PROGRAM PRG_Ladder
VAR
    bStart, bStop, bMotor, bButton, bClear, bLamp, bSkip, bRunning, bAlarm, bReady : BOOL;
    tonRun : TON;
    tElapsed : TIME;
END_VAR
VAR // added by the converter: edge detectors and wires of the graphical bodies
    _rt1 : R_TRIG;
END_VAR

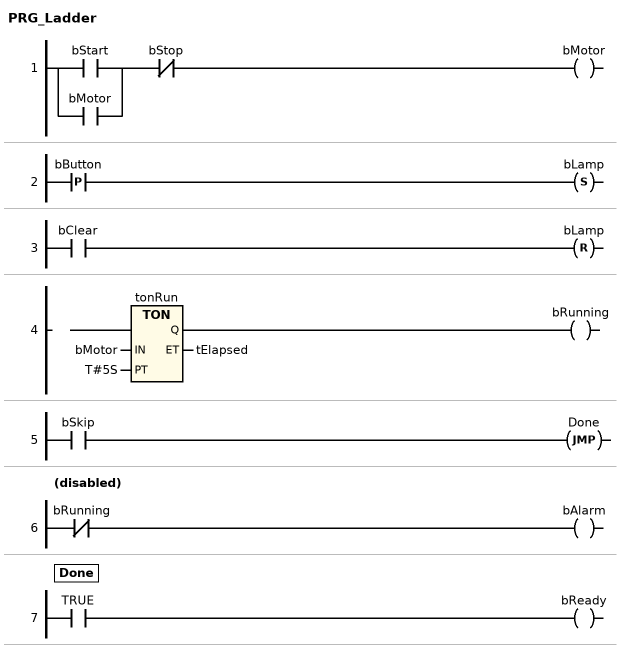
// NETWORK 1
bMotor := (bStart OR bMotor) AND NOT bStop;

// NETWORK 2
_rt1(CLK := bButton);
bLamp S= _rt1.Q;

// NETWORK 3
bLamp R= bClear;

// NETWORK 4
tonRun(IN := bMotor, PT := T#5S, ET => tElapsed); // TON
bRunning := tonRun.Q;

// NETWORK 5
IF bSkip THEN JMP Done; END_IF

// NETWORK 6 (disabled)
// bAlarm := NOT bRunning;

// NETWORK 7
Done:
bReady := TRUE;

END_PROGRAM

(* stored: Version 1.1.0.1, ProductVersion 3.1.4024.12
   POU PRG_Ladder: Id {00000000-0000-0000-0000-000000000001}, SpecialFunc None *)
